(* IEC 61131-3 sources: codesys-to-s7/tests/corpus/C2S7-POU-PRG/pos, 1 file *)

(* ---- input.st ---- *)
PROGRAM PRG_Case
VAR
    a : INT;
END_VAR
a := 1;
END_PROGRAM
